// TIA Portal project "EXERCICE2" (V16)

(* hardware
DEVICE "Station S7-1200_1"  S7-1200 Station
   slot 0: "Châssis_0"  S7-1200 Rack  Rack  V1.0
   slot 1: "PLC_1"  CPU 1214C AC/DC/Rly  6ES7 214-1BG40-0XB0  V4.4
DEVICE "HMI_1"  TP900 Comfort
   slot 0: "HMI_1"  TP900 Comfort  6AV2 124-0JC01-0AX0  16.0.0.0
   slot 1: "HMI_RT_1"  TP900 Comfort  6AV2 124-0JC01-0AX0  16.0.0.0
   slot 5: "HMI_1.IE_CP_1"  PROFINET Interface  16.0.0.0
      slot 1: "Interface PROFINET_1"  PROFINET Interface
         slot 1: "Port_1"  Port
         slot 2: "Port_2"  Port
   slot 7: "HMI_1.MPI/DP_CP_1"  MPI/DP Interface  16.0.0.0
*)

// ===== PLC "PLC_1"  CPU 1214C AC/DC/Rly =====

VAR_GLOBAL   // PLC tag table "Table de variables standard"
   "START" AT %I0.0 : Bool;
   "STOP" AT %I0.1 : Bool;
   "MOTEUR" AT %Q0.2 : Bool;
   "M" AT %M0.1 : Bool;
END_VAR

// folder: System blocks/Program resources

DATA_BLOCK "T1"   // DB1
{ S7_Optimized_Access := 'TRUE' }
AUTHOR : Simatic
FAMILY : IEC
NAME : IEC_TMR
VERSION : 1.0
// stored: InstanceOfName IEC_TIMER
"IEC_TIMER"
BEGIN
END_DATA_BLOCK

DATA_BLOCK "C1"   // DB2
{ S7_Optimized_Access := 'TRUE' }
AUTHOR : Simatic
FAMILY : IEC
NAME : CNTR
VERSION : 1.0
// stored: InstanceOfName IEC_COUNTER
"IEC_COUNTER"
BEGIN
END_DATA_BLOCK

// folder: (top level)

ORGANIZATION_BLOCK "Main"   // OB1, LAD, ProgramCycle
TITLE = "Main Program Sweep (Cycle)"
{ S7_Optimized_Access := 'TRUE' }
VERSION : 0.1
   VAR_INPUT
      Initial_Call : Bool;   // Initial call of this OB
      Remanence : Bool;   // =True, if remanent data are available
   END_VAR
BEGIN

REGION Network 1
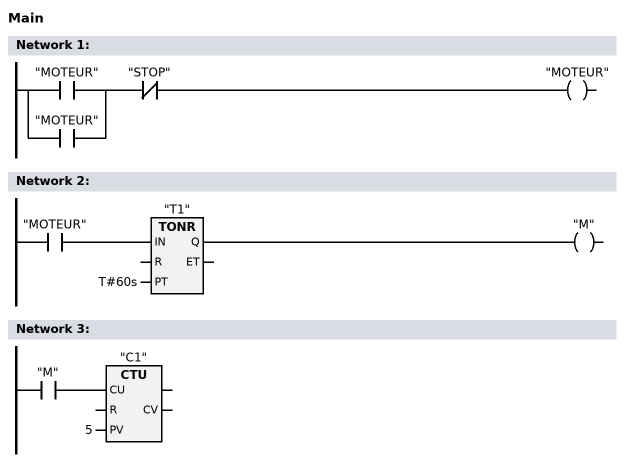
   RUNG wire#powerrail
      Contact( "MOTEUR" )
      wire#w1
      I_Contact( "STOP" )
      Coil( "MOTEUR" )
   END_RUNG
   RUNG wire#powerrail
      Contact( "MOTEUR" )
   END_RUNG wire#w1
   // the same network as SCL:
   "MOTEUR" := ("MOTEUR" OR "MOTEUR") AND NOT "STOP";
END_REGION

REGION Network 2
   "T1".TONR(IN := "MOTEUR", PT := T#60s);
   "M" := "T1".Q;
END_REGION

REGION Network 3
   "C1".CTU(CU := "M", PV := 5);
END_REGION
END_ORGANIZATION_BLOCK

(* ===== HMI "HMI_RT_1" =====
system functions are stored by id; their names below are inferred from use
connection "<Variabl>%": 

HMI tags "Table de variables standard"
   "Numéro_vue_variable" : UInt, internal
   "START_HMI" : Bool, 1 s
   "STOP_HMI" : UInt, internal
   "MOTEUR" : UInt, internal
   "4" : UInt, internal

text list "Nom_vue_liste_textes": 1 'Vue racine'

screen "Vue racine" 800x420, template "Modèle_1"
   on GenerateScreen: SetTag("Numéro_vue_variable", 1)
   Button "Bouton_1" at 15,13 size 144x80; TextOff 'START'
      on Press: SetBit("START_HMI")
      on Release: ResetBit("START_HMI")
   Button "Bouton_2" at 15,108 size 144x80; TextOff 'STOP'
      on Press: SetBit("STOP_HMI")
      on Release: ResetBit("STOP_HMI")
   Circle "Cercle_1" at 258,60 size 97x97
      Appearance <- "MOTEUR"
   TextField "Champ de texte_1" at 247,31 size 62x20; Text 'MOTEUR'

Template "Modèle_1" 800x420
   Button "Quitter" at 720,360 size 78x58; TextOff 'Quitter'; PictureOff "ExitRuntime_TP900_Comfort_TR"; PictureOn "ExitRuntime_TP900_Comfort_TR"
      on Release: StopRuntime(0)
   Button "Template_Button" at 640,360 size 78x58; TextOff 'Text'
   Button "Template_Button_1" at 560,360 size 78x58; TextOff 'Text'
   Button "Template_Button_2" at 480,360 size 78x58; TextOff 'Text'
   Button "Template_Button_3" at 400,360 size 78x58; TextOff 'Text'
   Button "Template_Button_4" at 321,360 size 78x58; TextOff 'Text'
   Button "Template_Button_5" at 241,360 size 78x58; TextOff 'Text'
   Button "Template_Button_6" at 161,360 size 78x58; TextOff 'Text'
   Button "Alarmes" at 81,360 size 78x58; TextOff 'Alarmes'; PictureOff "AlarmDisplay_TP900_Comfort_TR"; PictureOn "AlarmDisplay_TP900_Comfort_TR"
      on Release: function_ef3f5d25("Fenêtre des alarmes_non acquittée", -1)
   Button "Vue initiale" at 1,360 size 78x58; TextOff 'Vue initiale'; PictureOff "NavigateHome_TP900_Comfort_TR"; PictureOn "NavigateHome_TP900_Comfort_TR"
      on Release: ActivateScreen("Vue racine", 0)
*)